(* PLC project SelfHoldSample, CODESYS CODESYS V3.5 SP22 Patch 4 *)
(* stored: creationDateTime 2026-10-27T00:00:00, modificationDateTime 2026-10-27T00:00:00 *)

PROGRAM PLC_PRG

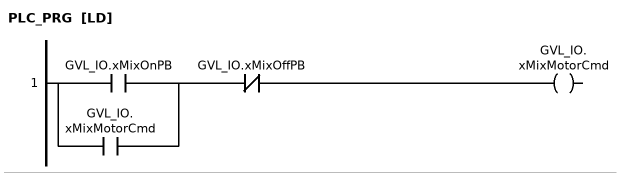
(* LD diagram, written out as Structured Text *)
(* 撹拌M 運転（自己保持） *)

GVL_IO.xMixMotorCmd := (GVL_IO.xMixOnPB OR GVL_IO.xMixMotorCmd) AND NOT GVL_IO.xMixOffPB;
END_PROGRAM
